TYPE ST_LimitOut :
STRUCT
	stP			: ST_Limit;	// kW
	stQ			: ST_Limit;	// kvar
	bResume		: BOOL;		// 출력 재개 중: 코어 램프가 재개 램프율을 쓴다
END_STRUCT
END_TYPE

(* stored: Version 1.1.0.1, ProductVersion 3.1.4024.15
   DUT ST_LimitOut: Id {7b9dc68f-cf87-4bd1-9b6a-3bc26306d5f6} *)
